// TIA Portal V18 export
VAR_GLOBAL   // PLC tag table "Default tag table"
   Forced_WO AT %I1500.0 : Bool;
   Trig_Buffer_ADIC AT %I1500.4 : Bool;
   Trig_Buffer_REMOV AT %I1500.5 : Bool;
   senor_filtro_oleo AT %I1000.0 : Bool;
   LEITOR_LEN AT %IB2283 : Byte;
   LEITURA_DONE AT %I2002.4 : Bool;
   sensor_vaselina AT %I1000.4 : Bool;
   Gatilho_ap_pneumaticaP105 AT %I221.6 : Bool;
   Sensor_RX1_RBX1 AT %I201.7 : Bool;
   Sensor_RX2_RBX2 AT %I201.6 : Bool;
   Sensor_cotovelo_mangueira AT %I1050.0 : Bool;
   Sensor_cotovelo AT %I1050.2 : Bool;
   Sensor_cotovelo_AD1600 AT %I1050.4 : Bool;
   Sensor_plug AT %I1050.6 : Bool;
   Tag_1 AT %QD1302 : DWord;
   Tag_2 AT %Q400.0 : Bool;
   Tag_3 AT %QW1310 : Int;
   SINAL_AP_SEMPRE_LIGADO AT %Q4000.0 : Bool;
   Tag_4 AT %QB1100 : Byte;
   RESET_DESOUTTER_P50 AT %Q8000.0 : Bool;
   RESET_DESOUTTER_P40 AT %Q6000.0 : Bool;
   Limpa_leitor AT %Q2000.7 : Bool;
   Buzzer_P01 AT %Q3.4 : Bool;
   Led_azul_P01 AT %Q3.2 : Bool;
   Led_red_P01 AT %Q3.0 : Bool;
   Led_verde_P01 AT %Q3.1 : Bool;
   Ledverde AT %Q1000.2 : Bool;
   Ledlaranja AT %Q1000.3 : Bool;
   LedVerde_vaselina AT %Q1000.6 : Bool;
   LedAmarelo_vaselina AT %Q1000.7 : Bool;
   LED_RX1_RBX1 AT %Q200.7 : Bool;
   LED_RX2_RBX2 AT %Q200.6 : Bool;
   Buzzer_P40 AT %Q5.4 : Bool;
   Led_azulP40 AT %Q5.2 : Bool;
   Led_VermelhoP40 AT %Q5.0 : Bool;
   Led_VerdeP40 AT %Q5.1 : Bool;
   Led_cotovelo_mangueira AT %Q1050.1 : Bool;
   Led_Cotovelo AT %Q1050.3 : Bool;
   Led_cotovelo_AD1600 AT %Q1050.5 : Bool;
   Led_Plug AT %Q1050.7 : Bool;
   FirstScan AT %M1.0 : Bool;
   DiagStatusUpdate AT %M1.1 : Bool;
   AlwaysTRUE AT %M1.2 : Bool;
   AlwaysFALSE AT %M1.3 : Bool;
   Clock_Byte AT %MB0 : Byte;
   Clock_10Hz AT %M0.0 : Bool;
   Clock_5Hz AT %M0.1 : Bool;
   "Clock_2.5Hz" AT %M0.2 : Bool;
   Clock_2Hz AT %M0.3 : Bool;
   "Clock_1.25Hz" AT %M0.4 : Bool;
   Clock_1Hz AT %M0.5 : Bool;
   "Clock_0.625Hz" AT %M0.6 : Bool;
   "Clock_0.5Hz" AT %M0.7 : Bool;
   status_10 AT %M1.4 : Bool;
   status_20 AT %M1.5 : Bool;
   status_40 AT %M1.6 : Bool;
   status_50 AT %M1.7 : Bool;
   status_60 AT %M6.0 : Bool;
   status_70 AT %M6.1 : Bool;
   status_80 AT %M6.2 : Bool;
   status_90 AT %M6.3 : Bool;
   status_100 AT %M6.4 : Bool;
   status_110 AT %M6.5 : Bool;
   status_120 AT %M6.6 : Bool;
   status_130 AT %M6.7 : Bool;
   BUSY AT %M7.6 : Bool;
   CYCLE_DONE_AREA_IHM AT %M8.0 : Bool;
   MODEZONE_DONE_AREA_IHM AT %M8.2 : Bool;
   CYCLE_DONE_IT_IHM AT %M8.4 : Bool;
   BOTAO_ACIONAR_MENSAGENS AT %M8.5 : Bool;
   Quantity_ok AT %MW10 : Int;
   BYPASSLEITOR AT %M7.7 : Bool;
   Inicia_apertadeiras AT %M4.4 : Bool;
   FORÇA_RECEITA_GERAL AT %M12.1 : Bool;
   CU_PRIMEIRO_POSTO AT %MW14 : Int;
   "POPID_INICO DE_LINHA" AT %M18.0 : LInt;
   Ready_to_copy AT %M2.0 : Bool;
   BYPASS_MOD_2 AT %M2.3 : Bool;
   BYPASS_MOD_1 AT %M2.4 : Bool;
   BYPASS_GERAL_EQUIP AT %M900.1 : Bool;
   "NOVO TESTE" AT %M9.5 : Bool;
   BYPASS_GERAL AT %M33.7 : Bool;
   ESVAZIAMENTO_FALCARE AT %M34.0 : Bool;
   ESVAZIA_FALCARE AT %M34.1 : Bool;
   ESVAZIA_MAIN_LINE AT %M34.2 : Bool;
   ESVAZIAMENTO_MAIN_LINE AT %M34.3 : Bool;
   ESVAZIA_FALCARE_1 AT %M34.4 : Bool;
   ESVAZIA_MAIN_LINE_1 AT %M34.5 : Bool;
   ERRO_ESVAZIAMENTO_LINHA AT %M34.6 : Bool;
   "CABINE EM MANUAL" AT %M34.7 : Bool;
   PRODUCAO_CONCLUIDA AT %M35.0 : Bool;
   GAP_E_EIXO_PENDURADO AT %M35.2 : Bool;
   VALIDACAO_EMERG_MOD1 AT %M35.3 : Bool;
   VALIDACAO_EMERG_MOD2 AT %M35.4 : Bool;
   "SINAL_DE RESET_GAP_CABINE" AT %M35.5 : Bool;
   BYPASS_TAMPA_CALIPER AT %M35.7 : Bool;
   INDEX_LEITOR AT %MW44 : UInt;
   CARACTER AT %MW46 : Int;
   RET_VAL AT %MW200 : Int;
   BYPASS_CABINE_EM_MODO_LOCAL AT %M42.5 : Bool;
   BYPASS_CAB_MODO_LOCAL AT %M42.6 : Bool;
   ACIONA_TELA AT %M43.1 : Bool;
   ERROR_COMUNICACAO_CABINE_SEND AT %M43.2 : Bool;
   ERROR_COMUNICACAO_CABINE_RECIVE AT %M43.3 : Bool;
   BYPASS_LEITURA AT %M43.4 : Bool;
   BORDA_MODZ1 AT %M43.5 : Bool;
   BYPASS_PY_JUNTA_RX_RBX AT %M43.6 : Bool;
   bypass_sem_receita AT %M2.7 : Bool;
   provisorio AT %M3.0 : Bool;
   BYPASS_PRENSA_LEMARB AT %M3.3 : Bool;
   TOOLRUNNING_POKA_JUNTA AT %M3.6 : Bool;
   BYPASS_TORQUIMETRO_DIGITAL AT %M4.2 : Bool;
   BYPASS_REULAGEM_ALAVANCA AT %M4.3 : Bool;
   ATIVA_FOR AT %M4.7 : Bool;
   PULSO_BY_P110 AT %M5.1 : Bool;
   set_modezone_done AT %M5.2 : Bool;
   giro_cabine AT %M5.3 : Bool;
   cabine_rodou AT %M5.4 : Bool;
   reset_md1 AT %M5.5 : Bool;
   reset_md2 AT %M5.6 : Bool;
   aux_gap AT %M7.0 : Bool;
   guarda_gap AT %M7.1 : Bool;
   chamada_forcada AT %MW16 : Int;
   Cabin_line_reference AT %M7.2 : Bool;
   SIGNAL_LOST_HELGE_2 AT %M8.6 : Bool;
   Habilita_matrix_P01 AT %M9.3 : Bool;
   Habilita_matrix_P05 AT %M9.4 : Bool;
   Habilita_matrix_P10 AT %M9.7 : Bool;
   Habilita_matrix_P15 AT %M26.0 : Bool;
   Habilita_matrix_P20 AT %M26.1 : Bool;
   Habilita_matrix_P30 AT %M26.2 : Bool;
   Habilita_matrix_P40 AT %M26.3 : Bool;
   Habilita_matrix_P50 AT %M26.4 : Bool;
   Habilita_matrix_P55 AT %M26.5 : Bool;
   Habilita_matrix_P60 AT %M26.6 : Bool;
   Habilita_matrix_P70 AT %M26.7 : Bool;
   Habilita_matrix_P75 AT %M27.0 : Bool;
   Habilita_matrix_P80 AT %M27.1 : Bool;
   Habilita_matrix_P90 AT %M27.2 : Bool;
   Habilita_matrix_P95 AT %M27.3 : Bool;
   Habilita_matrix_P100 AT %M27.4 : Bool;
   Habilita_matrix_P105 AT %M27.5 : Bool;
   Habilita_matrix_P110 AT %M27.6 : Bool;
   Habilita_matrix_P115 AT %M27.7 : Bool;
   Habilita_matrix_P120 AT %M42.7 : Bool;
   Habilita_matrix_P125 AT %M43.0 : Bool;
   Habilita_matrix_P130 AT %M56.0 : Bool;
   Habilita_matrix_P140 AT %M56.1 : Bool;
   Habilita_matrix_P150 AT %M56.2 : Bool;
   Habilita_matrix_QG AT %M56.3 : Bool;
   Bypass_graxa AT %M56.4 : Bool;
   Bypass_graxa_expedicao AT %M56.5 : Bool;
   JOBOK_PY_OLEO AT %M57.0 : Bool;
   antecipa_expedicao_1 AT %M57.1 : Bool;
   bahia AT %M58.1 : Bool;
   Count_gatilho AT %MW60 : Int;
END_VAR
VAR_GLOBAL CONSTANT   // user constants
   Config_OPC : Int := 17;
   maxConnectionsOPCUA : Int := 5;
END_VAR
